(* IEC 61131-3 sources: cia402-motion/templates, 1 file *)

(* ---- FB_Cia402Axis.st ---- *)
// FB_Cia402Axis and its types, as plain IEC 61131-3 Structured Text.
// The same declarations and body as the TwinCAT files beside it
// (FB_Cia402Axis.TcPOU and the four .TcDUT); tests/test_templates.py
// fails if the two drift apart. Reviewed and run against a simulated
// drive only: never compiled, never run on a real drive. Read
// templates/README.md first.

{attribute 'qualified_only'}
TYPE E_Cia402State :
(
    NotReadyToSwitchOn  := 0,
    SwitchOnDisabled    := 1,
    ReadyToSwitchOn     := 2,
    SwitchedOn          := 3,
    OperationEnabled    := 4,
    QuickStopActive     := 5,
    FaultReactionActive := 6,
    Fault               := 7,
    Unknown             := 8    // no state; or inputs that cannot be true
) INT;
END_TYPE

{attribute 'qualified_only'}
TYPE E_Cia402Step :
(
    Disabled        := 0,   // switched off, or on the way down
    WaitReady       := 10,  // T1: the drive leaves by itself
    Shutdown        := 11,  // T2: 0x0006
    SwitchOn        := 12,  // T3: 0x0007
    SetMode         := 13,  // 0x6060 written, 0x6061 awaited
    EnableOperation := 14,  // T4: 0x000F
    AbortEnable     := 15,  // bEnable fell during T4: 0x0007, wait
    Homing          := 20,  // controlword bit 4 held high
    Running         := 30,  // bValid: the set-points are the caller's
    ResetLow        := 40,  // bit 7 low, so that the next write is an edge
    ResetEdge       := 41,  // T15: 0x0080
    ResetRelease    := 42,  // bit 7 low again, after every attempt
    ResetPause      := 43,  // before the next attempt
    QuickStop       := 50,  // bQuickStop: 0x0002 held, then held down
    Error           := 90   // on the way down, waiting for bReset
) INT;
END_TYPE

TYPE ST_Cia402Drive :
STRUCT
    // Drive to PLC (TxPDO): copy in before each call. All three needed.
    nStatusword       : WORD;   // 0x6041
    nModesDisplay     : SINT;   // 0x6061
    nPositionActual   : DINT;   // 0x6064
    // PLC to drive (RxPDO): copy out after each call.
    nControlword      : WORD;   // 0x6040, written by the FB only
    nModesOfOperation : SINT;   // 0x6060, written by the FB only
    nTargetPosition   : DINT;   // 0x607A
    nTargetVelocity   : DINT;   // 0x60FF
    nTargetTorque     : INT;    // 0x6071
    // Caller to FB: controlword bits 4-6, 8, 9, sent only while bValid.
    nModeBits         : WORD;
END_STRUCT
END_TYPE

TYPE ST_Cia402Config :
STRUCT
    tStateTimeout     : TIME := T#2S;     // each transition, the mode switch
    tStopTimeout      : TIME := T#10S;    // a step down, a fault reaction
    tHomingTimeout    : TIME := T#60S;    // one whole homing run
    nResetAttempts    : UINT := 3;        // fault resets; 0 counts as 1
    tResetPause       : TIME := T#1S;     // between two reset attempts
    bQuickStopStays   : BOOL := FALSE;    // 0x605A is 5-8 on this drive
    nStandstillWindow : DINT := 0;        // position band, 0x6064 units
    tStandstill       : TIME := T#100MS;  // in the band this long: stopped
    tInputsInvalid    : TIME := T#100MS;  // bInputsValid FALSE this long: error
    bEnableAfterReset : BOOL := FALSE;    // TRUE: re-enable after bReset, as MC_Power
END_STRUCT
END_TYPE

FUNCTION_BLOCK FB_Cia402Axis
(*
    One CiA 402 drive: its state machine, the mode of operation, drive-based
    homing and fault reset. From the cia402-motion skill. It is a template:
    reviewed and run against a simulated drive, never compiled, never run
    on a real drive. Test it with reduced torque and speed limits before
    anyone stands near the machine. It is not a safety function: STO, SS1
    and safe stops belong in a safety controller.

    WHEN TO USE IT
    For a drive that makes the motion itself (PP, PV, PT, drive-based
    homing), or a PLC with no motion runtime. Where TwinCAT NC or CODESYS
    SoftMotion can drive the axis, use its axis and the MC_ blocks instead.
    Never both on one drive: both would write 0x6040.

    CONTRACT
    Call it once per cycle, unconditionally, in the task that exchanges the
    drive's process data. Copy 0x6041, 0x6061 and 0x6064 into stDrive
    before the call, in every mode, and stDrive's outputs to the drive
    after it.

    bEnable TRUE    Operation enabled in nMode. Once bValid is TRUE the
                    set-points in stDrive, and nModeBits, are yours.
                    Start a trajectory from where the FB left them: in
                    CSP, from stDrive.nTargetPosition.
    nMode = 6       Home with the method in 0x6098 (write it, and the
                    speeds, by SDO first). bValid then means homed. To
                    home again, drop bEnable or ask for another mode.
                    Change nMode at standstill only.
    bEnable FALSE   Stop and switch off: Disable operation (T5: 0x605C
                    decides how the motor stops), then T10. The same states
                    as cia402.py plan <state> sod, but T10 and T7 can go
                    out as 0x0002: see WHAT IT KEEPS TO.
    bReset          Rising edge: clear the error. If the drive is in
                    Fault, reset it first: bit 7 low, high, low. It does
                    not enable: after an error, bEnable must be FALSE once
                    before the FB enables again (stConfig.bEnableAfterReset
                    TRUE: it enables again with bEnable still TRUE).
    bQuickStop      TRUE: quick stop, from any step and over bEnable:
                    0x0002 held (T11: 0x605A decides how the motor stops).
                    One scan is enough. Not an error, and not a safety
                    function. A fault reset that has begun ends first, in
                    an error if it has to (16#8109), and 0x0002 goes out
                    then, so up to nResetAttempts limits later. The drive
                    goes to Switch on disabled and stays down until it is
                    there with bQuickStop and bEnable both FALSE, through
                    an error or a fault reset too, so that nothing
                    restarts it but a new bEnable. A drive that does not
                    take 0x0002 in tStateTimeout: 16#8108, and T5.
    bInputsValid    FALSE: this cycle's inputs are not the drive's (WcState,
                    the slave not in OP). Nothing is read and no step
                    changes; the outputs are held, but for bQuickStop.
                    Longer than tInputsInvalid: 16#8116. Default TRUE.

    Enabling always starts from Switch on disabled: a drive found anywhere
    else is taken down first, never taken over as it is. An error takes
    the drive down as bEnable FALSE does, and the FB stays down until
    bReset. It then stays down until bEnable has been FALSE, so that a
    reset never starts the axis. With stConfig.bEnableAfterReset it enables
    again while bEnable is still TRUE, as PLCopen MC_Power does after
    MC_Reset, unless a quick stop holds it down.
    nErrorID keeps the first error.

    WHAT IT KEEPS TO (the skill's references/state-machine.md)
    - One command at a time, held until the statusword shows the state it
      leads to, with a timeout. On the way up, any other state is an
      error. If bEnable falls while T4 may still be on its way, the FB
      sends 0x0007 and waits, so that a late T4 is stopped with T5. Only a
      quick stop cuts in: 0x0002 cannot be T9, whatever is on its way. If
      it falls while T2 or T3 may be, a new bEnable waits until the drive
      shows a new state, or for tStateTimeout: the Switch on disabled the
      FB sees may be older than the word.
    - Fault reset only from Fault: an edge on bit 7, released after every
      attempt, failed ones included. Never bit 7 with the enable bits.
    - Quick stop active is left only when the drive leaves it itself, or,
      where 0x605A keeps it there, at standstill. Never on a timer: that
      state is the stop ramp, and 0x0000 during it lets the motor coast.
    - On the way down, it never commands Operation enabled and never T9.
      The statusword is late, so a 0x000F already sent can have put the
      drive back there while the FB still sees Switched on. T10 and T7 go
      out as 0x0002, which is T11 there and not T9: 0x605A then decides how
      the motor stops, not 0x605C. Once bit 3 has been off for
      tStateTimeout no 0x000F can still come, and they go out as 0x0000,
      for a drive that does not take 0x0002.
    - One scan of a bad statusword does not send 0x0000, a fault reset or
      T2. A new state counts for those only if the next scan shows it too;
      until then the FB keeps bits 0-2 of its last word, or, while 0x000F
      may still land, sends 0x0002 as above. Fault and Fault reaction
      active add no 0x0000 of their own, until a reset. A bad word can
      still raise an error, and T11 or T5. A word that repeats is not told
      from the drive: see the README, What it cannot see.
    - Before T4 the set-points cannot move the motor: 0x607A = 0x6064,
      0x60FF = 0, 0x6071 = 0, bits 4-6, 8, 9 = 0. While the drive is
      enabled and they are not the caller's, the FB leaves them as they
      were, except that a mode switch makes the new mode's set-point safe
      a scan before it writes 0x6060. The mode counts once 0x6061 shows
      it.

    CHECK ON YOUR DRIVE (the skill's references/vendors/)
    - 0x605A 5-8 keeps the drive in Quick stop active at standstill, and
      any way down can end there, even with bQuickStop never used. Set
      stConfig.bQuickStopStays, and nStandstillWindow to the position
      jitter at standstill: the FB then leaves with T12 once the position
      has stayed in the band for tStandstill. Without the flag it waits
      for the drive to leave, which such a drive never does (safe, stuck).
    - Beckhoff's EL72x1 in DS402 reserves statusword bit 5. If it reads 0
      there, Ready to switch on and Switched on match no state, and the
      FB stops with 16#8115 after T2.
    - Beckhoff's EL72x1 in DS402 has no quick stop: controlword bit 2 is
      reserved there. LinMot's C125x-MI has no 0x605A. Try bQuickStop on
      such a drive before relying on it. If it ignores bit 2, a way down
      also waits in Ready to switch on until bit 3 has been off for
      tStateTimeout.
    - Statusword bit 12 in CSP is not checked: drives differ on it.
    - A homing result counts only after the drive has shown a phase with
      bits 12 and 13 both 0, from the scan bit 4 goes out on, so that an
      earlier run's result is not taken for this one. A drive that never
      shows one (an instant method 35 or 37 run twice) times out. Bit 13
      still set tStateTimeout after bit 4 went out is a homing error: a
      drive that refuses the method.
*)
VAR_INPUT
    bEnable      : BOOL;            // TRUE: run in nMode; FALSE: stop, off
    nMode        : SINT;            // 0x6060 code: 8 CSP, 1 PP, 6 homing...
    bReset       : BOOL;            // rising edge: clear, reset a fault
    bQuickStop   : BOOL;            // TRUE: T11, held. Not a safety stop
    bInputsValid : BOOL := TRUE;    // FALSE: the inputs are not the drive's
    stConfig     : ST_Cia402Config; // timeouts, reset retries, standstill
END_VAR
VAR_OUTPUT
    bValid      : BOOL;           // in nMode: the set-points are yours
    bBusy       : BOOL;           // on the way to what bEnable asks
    bError      : BOOL;
    nErrorID    : UDINT;          // 0 = none, else a cErr code below
    eDriveState : E_Cia402State;  // decoded from 0x6041
END_VAR
VAR_IN_OUT
    stDrive : ST_Cia402Drive;     // this axis' process data
END_VAR
VAR
    eStep            : E_Cia402Step := E_Cia402Step.Disabled;
    eStepPrev        : E_Cia402Step := E_Cia402Step.Disabled;
    eDrivePrev       : E_Cia402State := E_Cia402State.Unknown;
    fbResetTrig      : R_TRIG;
    fbStepTimer      : TON;       // the timeout of the step it is in
    fbStandstill     : TON;
    fbQuickStopTimer : TON;       // the drive has not taken 0x0002
    fbEnableWordOff  : TON;       // no 0x000F can still be on its way
    fbResetLimit     : TON;       // one attempt of a fault reset, at most
    fbUpWordOut      : TON;       // T2 or T3 can no longer come
    fbInputsInvalid  : TON;       // bInputsValid FALSE too long
    fbHomingStart    : TON;       // bit 4 out long enough to be taken
    tStepLimit       : TIME;
    bStepEntered     : BOOL;      // first scan in a new step
    bDriveMoved      : BOOL;      // the decoded state changed this scan
    bDriveSeen       : BOOL;      // the drive has left Not ready
    bAtRest          : BOOL;      // at rest, for a second scan
    bQuickStopHeld   : BOOL;      // asked for, not yet released
    bRestartHeld     : BOOL;      // an error: no enabling until bEnable FALSE
    bEnableNow       : BOOL;      // bEnable, unless an error holds it off
    bMoving          : BOOL;      // position left the standstill band
    nStandstillRef   : DINT;
    bHomingRunSeen   : BOOL;      // bits 12, 13 both 0 since bit 4
    bResetting       : BOOL;      // in one of the fault-reset steps
    bResetRequest    : BOOL;      // bReset rose while in Error
    bUpWordOut       : BOOL;      // T2 or T3 sent, not yet seen taken
    bSetModeLastScan : BOOL;      // last scan's outputs were SetMode's
    bRunningLastScan : BOOL;      // last scan's outputs were Running's
    nResetCount      : UINT;
END_VAR
VAR CONSTANT
    cModeBits       : WORD := 16#0370;   // controlword bits 4-6, 8, 9
    cResetSettle    : TIME := T#20MS;    // bit 7 low, before and after
    cErrNotReady    : UDINT := 16#8101;  // no Switch on disabled (T1)
    cErrShutdown    : UDINT := 16#8102;  // no Ready to switch on (T2)
    cErrSwitchOn    : UDINT := 16#8103;  // no Switched on (T3)
    cErrEnable      : UDINT := 16#8104;  // no Operation enabled (T4)
    cErrMode        : UDINT := 16#8105;  // 0x6061 never showed nMode
    cErrStop        : UDINT := 16#8106;  // did not get down in time
    cErrHomingTime  : UDINT := 16#8107;  // homing did not end in time
    cErrNoQuickStop : UDINT := 16#8108;  // drive did not take 0x0002
    cErrResetTime   : UDINT := 16#8109;  // fault reset did not end in time
    cErrDriveFault  : UDINT := 16#8110;  // drive in Fault: read 0x603F
    cErrResetFailed : UDINT := 16#8111;  // still in Fault after resets
    cErrQuickStop   : UDINT := 16#8112;  // Quick stop active, not ours
    cErrLeftState   : UDINT := 16#8113;  // drive moved where not asked
    cErrHoming      : UDINT := 16#8114;  // homing error, bit 13
    cErrStatusword  : UDINT := 16#8115;  // 0x6041 decodes to no state
    cErrInputs      : UDINT := 16#8116;  // bInputsValid FALSE too long
    cErrNoMode      : UDINT := 16#8120;  // nMode = 0
    cErrInvalidStep : UDINT := 16#8FFF;
END_VAR
// 0. bInputsValid FALSE: the inputs may not be the drive's (EtherCAT
//    WcState not 0 or the slave not in OP, a CANopen PDO not received).
//    Nothing is read from them and no step changes: every output stays as
//    the last scan left it, 0x6040 included, but for a quick stop asked
//    for, which sends 0x0002. The timers run on, so a step judged on the
//    first valid scan has had the time that passed. Longer than
//    tInputsInvalid is an error, and the last word still goes out until
//    the inputs are valid again: the drive's own reaction to a lost bus
//    (0x6007) is what stops it then.
fbInputsInvalid(IN := NOT bInputsValid, PT := stConfig.tInputsInvalid);
IF NOT bInputsValid THEN
    IF bQuickStop THEN
        bQuickStopHeld := TRUE;
    END_IF
    IF bQuickStopHeld AND NOT bResetting AND NOT fbQuickStopTimer.Q THEN
        stDrive.nControlword := 16#0002;
    END_IF
    IF fbInputsInvalid.Q AND (eStep <> E_Cia402Step.Error) THEN
        nErrorID := cErrInputs;
        eStep    := E_Cia402Step.Error;
    END_IF
    bValid := (eStep = E_Cia402Step.Running) AND NOT bQuickStopHeld;
    bError := (eStep = E_Cia402Step.Error);
    bBusy  := bBusy AND NOT bError;
ELSE
    // 1. Decode 0x6041. Each state has its own mask: bit 5 belongs to four of
    //    them and is a don't-care in the other four. A word that matches none
    //    is read fault-first, as cia402.py decode sw does.
    IF (stDrive.nStatusword AND 16#004F) = 16#0000 THEN
        eDriveState := E_Cia402State.NotReadyToSwitchOn;
    ELSIF (stDrive.nStatusword AND 16#004F) = 16#0040 THEN
        eDriveState := E_Cia402State.SwitchOnDisabled;
    ELSIF (stDrive.nStatusword AND 16#006F) = 16#0021 THEN
        eDriveState := E_Cia402State.ReadyToSwitchOn;
    ELSIF (stDrive.nStatusword AND 16#006F) = 16#0023 THEN
        eDriveState := E_Cia402State.SwitchedOn;
    ELSIF (stDrive.nStatusword AND 16#006F) = 16#0027 THEN
        eDriveState := E_Cia402State.OperationEnabled;
    ELSIF (stDrive.nStatusword AND 16#006F) = 16#0007 THEN
        eDriveState := E_Cia402State.QuickStopActive;
    ELSIF (stDrive.nStatusword AND 16#0008) = 0 THEN
        eDriveState := E_Cia402State.Unknown;
    ELSIF (stDrive.nStatusword AND 16#0007) = 16#0007 THEN
        eDriveState := E_Cia402State.FaultReactionActive;
    ELSE
        eDriveState := E_Cia402State.Fault;
    END_IF

    // A drive never goes back to Not ready to switch on. Seen after another
    // state, that word means the inputs are not the drive's: a bus restart, a
    // copy that never happened. 0x0000 sent then could be T9.
    IF (eDriveState <> E_Cia402State.NotReadyToSwitchOn)
       AND (eDriveState <> E_Cia402State.Unknown)
    THEN
        bDriveSeen := TRUE;
    ELSIF bDriveSeen AND (eDriveState = E_Cia402State.NotReadyToSwitchOn) THEN
        eDriveState := E_Cia402State.Unknown;
    END_IF

    // 2. Every block that carries state is called here, once per scan, above
    //    the state machine that reads it.
    fbResetTrig(CLK := bReset);

    bStepEntered := (eStep <> eStepPrev);
    bDriveMoved  := (eDriveState <> eDrivePrev);
    eStepPrev    := eStep;
    eDrivePrev   := eDriveState;

    // At rest only from the second scan: one bad word is no reason to send
    // 0x0000, or to let a quick stop go.
    bAtRest := NOT bDriveMoved
               AND ((eDriveState = E_Cia402State.SwitchOnDisabled)
                    OR (eDriveState = E_Cia402State.NotReadyToSwitchOn));

    bResetting := (eStep = E_Cia402Step.ResetLow)
                  OR (eStep = E_Cia402Step.ResetEdge)
                  OR (eStep = E_Cia402Step.ResetRelease)
                  OR (eStep = E_Cia402Step.ResetPause);

    // A reset asked for in Error is kept until it can be acted on, so that an
    // edge in Fault reaction active is not lost.
    IF eStep <> E_Cia402Step.Error THEN
        bResetRequest := FALSE;
    ELSIF fbResetTrig.Q THEN
        bResetRequest := TRUE;
    END_IF

    // After an error the axis enables again only on a bEnable that was FALSE
    // once the error had been cleared: a reset must not start it. A bEnable
    // that falls and rises during the error does not count.
    IF (eStep = E_Cia402Step.Error) AND NOT stConfig.bEnableAfterReset THEN
        bRestartHeld := TRUE;
    ELSIF NOT bEnable OR stConfig.bEnableAfterReset THEN
        bRestartHeld := FALSE;
    END_IF
    bEnableNow := bEnable AND NOT bRestartHeld;

    // The timeout of the step the FB is in. IN low on the scan the step or
    // the drive's state changed re-arms it, so every transition gets a full
    // timeout of its own.
    CASE eStep OF
        E_Cia402Step.Homing:
            tStepLimit := stConfig.tHomingTimeout;
        E_Cia402Step.Disabled, E_Cia402Step.Error:
            tStepLimit := stConfig.tStopTimeout;
        E_Cia402Step.ResetLow, E_Cia402Step.ResetRelease:
            tStepLimit := cResetSettle;
        E_Cia402Step.ResetPause:
            tStepLimit := stConfig.tResetPause;
    ELSE
        tStepLimit := stConfig.tStateTimeout;
    END_CASE
    fbStepTimer(IN := NOT (bStepEntered OR bDriveMoved), PT := tStepLimit);

    // Standstill, for leaving Quick stop active where 0x605A keeps the drive
    // there: the position has stayed inside the band for tStandstill. It
    // measures the motor, not the time since the stop began.
    bMoving := ABS(stDrive.nPositionActual - nStandstillRef)
               > stConfig.nStandstillWindow;
    IF bMoving THEN
        nStandstillRef := stDrive.nPositionActual;
    END_IF
    fbStandstill(IN := stConfig.bQuickStopStays
                       AND (eDriveState = E_Cia402State.QuickStopActive)
                       AND NOT bMoving,
                 PT := stConfig.tStandstill);

    // A quick stop is kept, through an error or a fault reset too, until the
    // drive is down with bQuickStop and bEnable both FALSE: only a new
    // bEnable restarts the axis. The timer gives the drive tStateTimeout to
    // take 0x0002. It never runs in Quick stop active: that state is the stop
    // ramp. Nor in a fault reset: 0x0002 has not gone out yet.
    IF bQuickStop THEN
        bQuickStopHeld := TRUE;
    ELSIF bAtRest AND NOT bEnable THEN
        bQuickStopHeld := FALSE;
    END_IF
    fbQuickStopTimer(IN := bQuickStopHeld AND NOT bAtRest
                           AND (eDriveState <> E_Cia402State.QuickStopActive)
                           AND NOT bResetting,
                     PT := stConfig.tStateTimeout);

    // How long the FB's own words have been without bit 3. It reads no state: a
    // statusword that flips between two states must not re-arm it.
    fbEnableWordOff(IN := (stDrive.nControlword AND 16#0008) = 0,
                    PT := stConfig.tStateTimeout);

    // A fault reset ends, whatever the drive shows: fbStepTimer waits out
    // Fault reaction active with no limit, and a state change re-arms it. This
    // limit is re-armed only by the attempt counted on the way into
    // ResetPause, and the attempts run out. It allows one attempt whole, with
    // its pause, and a fault reaction as long as a stop; the second
    // tStateTimeout is for the scans each step loses, and the statusword's lag.
    fbResetLimit(IN := bResetting
                       AND NOT (bStepEntered
                                AND (eStep = E_Cia402Step.ResetPause)),
                 PT := stConfig.tResetPause + stConfig.tStateTimeout
                       + stConfig.tStateTimeout + stConfig.tStopTimeout);

    // A 0x0006 or 0x0007 left behind when bEnable fell has been taken, or
    // ignored, once the drive shows a new state, or after tStateTimeout. Until
    // then the Switch on disabled the FB sees may be older than that word.
    fbUpWordOut(IN := bUpWordOut, PT := stConfig.tStateTimeout);
    IF bDriveMoved OR fbUpWordOut.Q THEN
        bUpWordOut := FALSE;
    END_IF

    // Homing, statusword bits 13, 12, 10. Bits 12 and 13 both 0 (in progress,
    // or not started) cannot be left over from an earlier run. Outside homing
    // this follows the latest phase; in it, it latches. A drive that
    // refuses the start sets bit 13 without such a phase, and bit 13 left
    // from an earlier run then never clears: still there tStateTimeout after
    // bit 4 went out, it is this run's.
    IF (stDrive.nStatusword AND 16#3000) = 0 THEN
        bHomingRunSeen := TRUE;
    ELSIF eStep <> E_Cia402Step.Homing THEN
        bHomingRunSeen := FALSE;
    END_IF
    fbHomingStart(IN := (eStep = E_Cia402Step.Homing),
                  PT := stConfig.tStateTimeout);

    // 3. A statusword that decodes to no state is an error in every step; a
    //    fault is one in every step but the reset itself. A quick stop takes
    //    over from every step but Error and the reset, which ends first.
    IF eStep <> E_Cia402Step.Error THEN
        IF eDriveState = E_Cia402State.Unknown THEN
            nErrorID := cErrStatusword;
            eStep    := E_Cia402Step.Error;
        ELSIF NOT bResetting
              AND ((eDriveState = E_Cia402State.Fault)
                   OR (eDriveState = E_Cia402State.FaultReactionActive))
        THEN
            nErrorID := cErrDriveFault;
            eStep    := E_Cia402Step.Error;
        ELSIF bResetting AND fbResetLimit.Q THEN
            nErrorID := cErrResetTime;
            eStep    := E_Cia402Step.Error;
        ELSIF bQuickStopHeld AND NOT bResetting THEN
            eStep := E_Cia402Step.QuickStop;
        END_IF
    END_IF

    // 4. Transitions. Each step names the state it waits for and the state it
    //    may still be in; anything else, or its timeout, is an error.
    CASE eStep OF

        E_Cia402Step.Disabled:
            // On the way down (outputs below). Enabling starts only from
            // Switch on disabled, where no command of the way down can still
            // be on its way.
            IF bEnableNow AND nMode = 0 THEN
                nErrorID := cErrNoMode;
                eStep    := E_Cia402Step.Error;
            ELSIF bEnableNow
                  AND eDriveState = E_Cia402State.NotReadyToSwitchOn
            THEN
                eStep := E_Cia402Step.WaitReady;
            ELSIF bEnableNow AND NOT bDriveMoved AND NOT bUpWordOut
                  AND eDriveState = E_Cia402State.SwitchOnDisabled
            THEN
                eStep := E_Cia402Step.Shutdown;
            ELSIF fbStepTimer.Q
                  AND ((eDriveState = E_Cia402State.OperationEnabled)
                       OR (eDriveState = E_Cia402State.SwitchedOn)
                       OR (eDriveState = E_Cia402State.ReadyToSwitchOn))
            THEN
                nErrorID := cErrStop;
                eStep    := E_Cia402Step.Error;
            END_IF

        E_Cia402Step.WaitReady:
            IF NOT bEnable THEN
                eStep := E_Cia402Step.Disabled;
            ELSIF eDriveState = E_Cia402State.SwitchOnDisabled THEN
                eStep := E_Cia402Step.Shutdown;
            ELSIF eDriveState <> E_Cia402State.NotReadyToSwitchOn THEN
                nErrorID := cErrLeftState;
                eStep    := E_Cia402Step.Error;
            ELSIF fbStepTimer.Q THEN
                nErrorID := cErrNotReady;
                eStep    := E_Cia402Step.Error;
            END_IF

        E_Cia402Step.Shutdown:
            IF NOT bEnable THEN
                bUpWordOut := TRUE;
                eStep      := E_Cia402Step.Disabled;
            ELSIF eDriveState = E_Cia402State.ReadyToSwitchOn THEN
                eStep := E_Cia402Step.SwitchOn;
            ELSIF eDriveState <> E_Cia402State.SwitchOnDisabled THEN
                nErrorID := cErrLeftState;
                eStep    := E_Cia402Step.Error;
            ELSIF fbStepTimer.Q THEN
                nErrorID := cErrShutdown;
                eStep    := E_Cia402Step.Error;
            END_IF

        E_Cia402Step.SwitchOn:
            IF NOT bEnable THEN
                bUpWordOut := TRUE;
                eStep      := E_Cia402Step.Disabled;
            ELSIF eDriveState = E_Cia402State.SwitchedOn THEN
                eStep := E_Cia402Step.SetMode;
            ELSIF eDriveState <> E_Cia402State.ReadyToSwitchOn THEN
                nErrorID := cErrLeftState;
                eStep    := E_Cia402Step.Error;
            ELSIF fbStepTimer.Q THEN
                nErrorID := cErrSwitchOn;
                eStep    := E_Cia402Step.Error;
            END_IF

        E_Cia402Step.SetMode:
            // In Switched on on the way up, in Operation enabled when the mode
            // changes while running; the drive must stay where it was. Done
            // once 0x6060 has gone out as nMode and 0x6061 shows it.
            IF NOT bEnable THEN
                eStep := E_Cia402Step.Disabled;
            ELSIF nMode = 0 THEN
                nErrorID := cErrNoMode;
                eStep    := E_Cia402Step.Error;
            ELSIF eDriveState = E_Cia402State.QuickStopActive THEN
                nErrorID := cErrQuickStop;
                eStep    := E_Cia402Step.Error;
            ELSIF bDriveMoved
                  OR ((eDriveState <> E_Cia402State.SwitchedOn)
                      AND (eDriveState <> E_Cia402State.OperationEnabled))
            THEN
                nErrorID := cErrLeftState;
                eStep    := E_Cia402Step.Error;
            ELSIF (stDrive.nModesOfOperation = nMode)
                  AND (stDrive.nModesDisplay = nMode)
            THEN
                IF eDriveState = E_Cia402State.SwitchedOn THEN
                    eStep := E_Cia402Step.EnableOperation;
                ELSIF nMode = 6 THEN
                    eStep := E_Cia402Step.Homing;
                ELSE
                    eStep := E_Cia402Step.Running;
                END_IF
            ELSIF fbStepTimer.Q THEN
                nErrorID := cErrMode;
                eStep    := E_Cia402Step.Error;
            END_IF

        E_Cia402Step.EnableOperation:
            IF eDriveState = E_Cia402State.OperationEnabled THEN
                IF NOT bEnable THEN
                    eStep := E_Cia402Step.Disabled;
                ELSIF (nMode <> stDrive.nModesOfOperation)
                      OR (nMode <> stDrive.nModesDisplay)
                THEN
                    eStep := E_Cia402Step.SetMode;
                ELSIF nMode = 6 THEN
                    eStep := E_Cia402Step.Homing;
                ELSE
                    eStep := E_Cia402Step.Running;
                END_IF
            ELSIF eDriveState <> E_Cia402State.SwitchedOn THEN
                nErrorID := cErrLeftState;
                eStep    := E_Cia402Step.Error;
            ELSIF NOT bEnable THEN
                eStep := E_Cia402Step.AbortEnable;
            ELSIF fbStepTimer.Q THEN
                nErrorID := cErrEnable;
                eStep    := E_Cia402Step.Error;
            END_IF

        E_Cia402Step.AbortEnable:
            // 0x000F may still be on its way, and bEnable FALSE stops with T5,
            // not T11. 0x0007 is T5 in Operation enabled and nothing in
            // Switched on; after tStateTimeout there no T4 can still come.
            IF (eDriveState <> E_Cia402State.SwitchedOn) OR fbStepTimer.Q THEN
                eStep := E_Cia402Step.Disabled;
            END_IF

        E_Cia402Step.Homing:
            // Dropping bit 4 interrupts the run: bEnable FALSE and a mode
            // change both do that, through the outputs of the next step.
            IF NOT bEnable THEN
                eStep := E_Cia402Step.Disabled;
            ELSIF eDriveState = E_Cia402State.QuickStopActive THEN
                nErrorID := cErrQuickStop;
                eStep    := E_Cia402Step.Error;
            ELSIF eDriveState <> E_Cia402State.OperationEnabled THEN
                nErrorID := cErrLeftState;
                eStep    := E_Cia402Step.Error;
            ELSIF (nMode <> stDrive.nModesOfOperation)
                  OR (nMode <> stDrive.nModesDisplay)
            THEN
                eStep := E_Cia402Step.SetMode;
            ELSIF (bHomingRunSeen OR fbHomingStart.Q)
                  AND ((stDrive.nStatusword AND 16#2000) <> 0)
            THEN
                nErrorID := cErrHoming;
                eStep    := E_Cia402Step.Error;
            ELSIF bHomingRunSeen
                  AND ((stDrive.nStatusword AND 16#3400) = 16#1400)
            THEN
                eStep := E_Cia402Step.Running;
            ELSIF fbStepTimer.Q THEN
                nErrorID := cErrHomingTime;
                eStep    := E_Cia402Step.Error;
            END_IF

        E_Cia402Step.Running:
            IF NOT bEnable THEN
                eStep := E_Cia402Step.Disabled;
            ELSIF eDriveState = E_Cia402State.QuickStopActive THEN
                nErrorID := cErrQuickStop;
                eStep    := E_Cia402Step.Error;
            ELSIF eDriveState <> E_Cia402State.OperationEnabled THEN
                nErrorID := cErrLeftState;
                eStep    := E_Cia402Step.Error;
            ELSIF (nMode <> stDrive.nModesOfOperation)
                  OR (nMode <> stDrive.nModesDisplay)
            THEN
                eStep := E_Cia402Step.SetMode;
            END_IF

        E_Cia402Step.ResetLow, E_Cia402Step.ResetPause:
            // A drive can leave Fault without this edge: a reset it took late,
            // its own input. Bit 7 is low already, so a state that has lasted
            // the whole step is judged here, and no attempt is counted: none
            // was made. Fault reaction active is still the fault: it is waited
            // for, up to fbResetLimit.
            IF fbStepTimer.Q THEN
                IF eDriveState = E_Cia402State.Fault THEN
                    eStep := E_Cia402Step.ResetEdge;
                ELSIF eDriveState = E_Cia402State.SwitchOnDisabled THEN
                    nErrorID := 0;
                    eStep    := E_Cia402Step.Disabled;
                ELSIF eDriveState <> E_Cia402State.FaultReactionActive THEN
                    nErrorID := cErrLeftState;
                    eStep    := E_Cia402Step.Error;
                END_IF
            END_IF

        E_Cia402Step.ResetEdge:
            // Hold the edge until the drive leaves Fault or the timeout, then
            // release bit 7 either way. A state seen for one scan may be a bad
            // word: the step stays, so that the drive still gets its edge.
            IF ((eDriveState <> E_Cia402State.Fault) AND NOT bDriveMoved)
               OR fbStepTimer.Q
            THEN
                eStep := E_Cia402Step.ResetRelease;
            END_IF

        E_Cia402Step.ResetRelease:
            IF fbStepTimer.Q THEN
                IF eDriveState = E_Cia402State.SwitchOnDisabled THEN
                    nErrorID := 0;
                    eStep    := E_Cia402Step.Disabled;
                ELSIF (eDriveState <> E_Cia402State.Fault)
                      AND (eDriveState <> E_Cia402State.FaultReactionActive)
                THEN
                    nErrorID := cErrLeftState;
                    eStep    := E_Cia402Step.Error;
                ELSE
                    // Still faulted: the cause is still there. Read 0x603F.
                    nResetCount := nResetCount + 1;
                    IF nResetCount < stConfig.nResetAttempts THEN
                        eStep := E_Cia402Step.ResetPause;
                    ELSE
                        nErrorID := cErrResetFailed;
                        eStep    := E_Cia402Step.Error;
                    END_IF
                END_IF
            END_IF

        E_Cia402Step.QuickStop:
            IF NOT bQuickStopHeld THEN
                eStep := E_Cia402Step.Disabled;
            ELSIF fbQuickStopTimer.Q THEN
                nErrorID := cErrNoQuickStop;
                eStep    := E_Cia402Step.Error;
            END_IF

        E_Cia402Step.Error:
            // On the way down, as Disabled. A reset waits while the drive is
            // in Fault reaction active or its statusword decodes to nothing,
            // and for a second scan of a new state: ResetLow sends 0x0000.
            IF bResetRequest AND NOT bDriveMoved THEN
                IF eDriveState = E_Cia402State.Fault THEN
                    nErrorID    := 0;
                    nResetCount := 0;
                    eStep       := E_Cia402Step.ResetLow;
                ELSIF (eDriveState <> E_Cia402State.FaultReactionActive)
                      AND (eDriveState <> E_Cia402State.Unknown)
                THEN
                    nErrorID := 0;
                    eStep    := E_Cia402Step.Disabled;
                END_IF
            END_IF

    ELSE
        nErrorID := cErrInvalidStep;
        eStep    := E_Cia402Step.Error;
    END_CASE

    // 5. Outputs, from the step the FB is in after this scan's transitions:
    //    the word sent always belongs to the step that holds it.
    CASE eStep OF

        E_Cia402Step.Disabled, E_Cia402Step.Error:
            // The way down: the states of cia402.py plan <state> sod, with
            // 0x0002 for T7, T10 while 0x000F may still come. One word per
            // state, but for the first scan of a state: see bDriveMoved below.
            CASE eDriveState OF
                E_Cia402State.OperationEnabled:
                    // 0x0002 sent below may have gone out after a statusword
                    // that is only now showing the climb: hold it, one command
                    // at a time, until no 0x000F can still come.
                    IF (bQuickStopHeld AND NOT fbQuickStopTimer.Q)
                       OR ((stDrive.nControlword = 16#0002)
                           AND NOT fbEnableWordOff.Q)
                    THEN
                        stDrive.nControlword := 16#0002;   // T11, in Error
                    ELSE
                        stDrive.nControlword := 16#0007;   // T5, per 0x605C
                    END_IF
                E_Cia402State.QuickStopActive:
                    IF fbStandstill.Q THEN
                        stDrive.nControlword := 16#0000;   // T12, stopped
                    ELSE
                        stDrive.nControlword := 16#0002;   // let it finish
                    END_IF
                E_Cia402State.SwitchedOn, E_Cia402State.ReadyToSwitchOn:
                    // T10, T7. 0x0002 leaves these two as 0x0000 does, but a
                    // late statusword may hide a 0x000F that has put the drive
                    // back in Operation enabled: there it is T11, and 0x0000
                    // is T9. A drive may ignore bit 2 and read it as Shutdown.
                    // Once bit 3 has been off for tStateTimeout no 0x000F can
                    // still come. Seen for one scan it may be a bad word: keep
                    // the last word, never 0x0002 here, which would chase
                    // 0x0000 on such a drive.
                    IF fbEnableWordOff.Q AND NOT bDriveMoved THEN
                        stDrive.nControlword := 16#0000;
                    ELSIF fbEnableWordOff.Q THEN
                        stDrive.nControlword := stDrive.nControlword
                                                AND 16#0007;
                    ELSE
                        stDrive.nControlword := 16#0002;
                    END_IF
                E_Cia402State.Fault, E_Cia402State.FaultReactionActive,
                E_Cia402State.Unknown:
                    // Keep the last word, less enable operation, the mode bits
                    // and bit 7: it cannot enable, and it cannot cut power. A
                    // drive in Fault ignores it, and the word may be a bad one.
                    IF bQuickStopHeld AND NOT fbQuickStopTimer.Q THEN
                        stDrive.nControlword := 16#0002;
                    ELSE
                        stDrive.nControlword := stDrive.nControlword
                                                AND 16#0007;
                    END_IF
            ELSE
                // At rest. Seen for one scan it may be a bad word: to a drive
                // still enabled, 0x0000 would be T9.
                IF bDriveMoved THEN
                    stDrive.nControlword := stDrive.nControlword AND 16#0007;
                ELSE
                    stDrive.nControlword := 16#0000;
                END_IF
            END_CASE

        E_Cia402Step.WaitReady, E_Cia402Step.ResetLow,
        E_Cia402Step.ResetRelease, E_Cia402Step.ResetPause:
            stDrive.nControlword := 16#0000;

        E_Cia402Step.Shutdown:
            stDrive.nControlword := 16#0006;   // T2

        E_Cia402Step.SwitchOn, E_Cia402Step.AbortEnable:
            stDrive.nControlword := 16#0007;   // T3; or T5 after a late T4

        E_Cia402Step.SetMode:
            IF eDriveState = E_Cia402State.OperationEnabled THEN
                stDrive.nControlword := 16#000F;   // hold Operation enabled
            ELSE
                stDrive.nControlword := 16#0007;   // hold Switched on
            END_IF
            IF bSetModeLastScan THEN
                stDrive.nModesOfOperation := nMode;
            END_IF

        E_Cia402Step.EnableOperation:
            stDrive.nControlword := 16#000F;   // T4

        E_Cia402Step.Homing:
            stDrive.nControlword := 16#001F;   // bit 4: homing start, held

        E_Cia402Step.Running:
            // The caller's bits from the second scan on: on the first, the
            // caller has not seen bValid yet.
            IF (nMode = 6) OR NOT bRunningLastScan THEN
                stDrive.nControlword := 16#000F;
            ELSE
                stDrive.nControlword := 16#000F
                                        OR (stDrive.nModeBits AND cModeBits);
            END_IF

        E_Cia402Step.QuickStop:
            // 0x0002 is T11 in Operation enabled and goes to Switch on disabled
            // from the two states below it, so that a T4 still on its way meets
            // T11. 0x0000 there could be T9.
            IF bAtRest OR fbStandstill.Q THEN
                stDrive.nControlword := 16#0000;   // at rest; or T12, stopped
            ELSE
                stDrive.nControlword := 16#0002;   // T11, held
            END_IF

        E_Cia402Step.ResetEdge:
            // T15, a rising edge on bit 7: only ever sent to a drive in Fault.
            IF eDriveState = E_Cia402State.Fault THEN
                stDrive.nControlword := 16#0080;
            ELSE
                stDrive.nControlword := 16#0000;
            END_IF

    ELSE
        stDrive.nControlword := 16#0000;
    END_CASE
    bSetModeLastScan := (eStep = E_Cia402Step.SetMode);
    bRunningLastScan := (eStep = E_Cia402Step.Running);

    // 6. Set-points. From bValid on they are the caller's. Without torque the
    //    FB holds them where enabling cannot move the motor. With the drive
    //    enabled it leaves them as they were, so that it never steps one the
    //    drive is following; a mode switch makes the new mode's set-point
    //    safe. The caller's mode bits are cleared until bValid. One scan of
    //    a new state does not count: the drive may still be following.
    IF (eStep = E_Cia402Step.Running)
       OR (bDriveMoved AND (eStep <> E_Cia402Step.SetMode))
    THEN
        ;
    ELSIF (eDriveState <> E_Cia402State.OperationEnabled)
          AND (eDriveState <> E_Cia402State.QuickStopActive)
    THEN
        stDrive.nTargetPosition := stDrive.nPositionActual;
        stDrive.nTargetVelocity := 0;
        stDrive.nTargetTorque   := 0;
        stDrive.nModeBits       := 0;
    ELSE
        IF eStep = E_Cia402Step.SetMode THEN
            CASE nMode OF
                1, 8:
                    stDrive.nTargetPosition := stDrive.nPositionActual;
                3, 9:
                    stDrive.nTargetVelocity := 0;
                4, 10, 11:
                    stDrive.nTargetTorque := 0;
            ELSE
                ;   // a mode of the drive's own: see its manual
            END_CASE
        END_IF
        stDrive.nModeBits := 0;
    END_IF

    bValid := (eStep = E_Cia402Step.Running);
    bError := (eStep = E_Cia402Step.Error);
    bBusy  := NOT bValid AND NOT bError
              AND ((bEnableNow AND (eStep <> E_Cia402Step.QuickStop))
                   OR NOT bAtRest);
END_IF
END_FUNCTION_BLOCK
